Omron CX-Programmer project OmronTeachingExample (CX-Programmer 9.73)

# PLC ExamplePLC: CP1H XA

## Program Main (cyclic task 0)

### Section Section1

### Section Analog_Validity

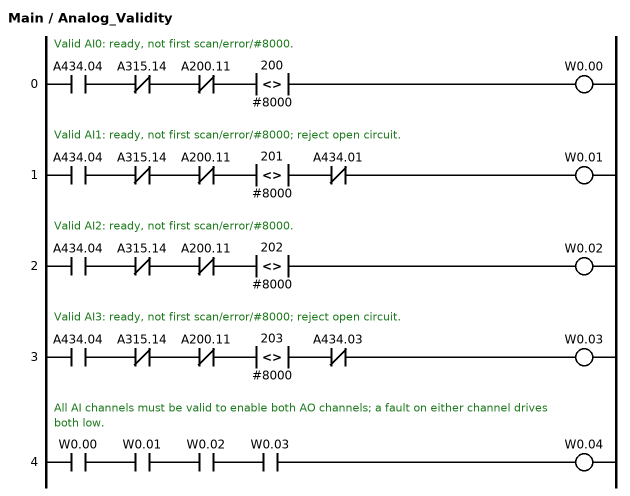
; rung 0: Valid AI0: ready, not first scan/error/#8000.
LD A434.04
ANDNOT A315.14
ANDNOT A200.11
AND<>(305) 200 #8000
OUT W0.00
; rung 1: Valid AI1: ready, not first scan/error/#8000; reject open circuit.
LD A434.04
ANDNOT A315.14
ANDNOT A200.11
AND<>(305) 201 #8000
ANDNOT A434.01
OUT W0.01
; rung 2: Valid AI2: ready, not first scan/error/#8000.
LD A434.04
ANDNOT A315.14
ANDNOT A200.11
AND<>(305) 202 #8000
OUT W0.02
; rung 3: Valid AI3: ready, not first scan/error/#8000; reject open circuit.
LD A434.04
ANDNOT A315.14
ANDNOT A200.11
AND<>(305) 203 #8000
ANDNOT A434.03
OUT W0.03
; rung 4: All AI channels must be valid to enable both AO channels; a fault on either channel drives both low.
LD W0.00
AND W0.01
AND W0.02
AND W0.03
OUT W0.04

### Section HMI_Input_Publication

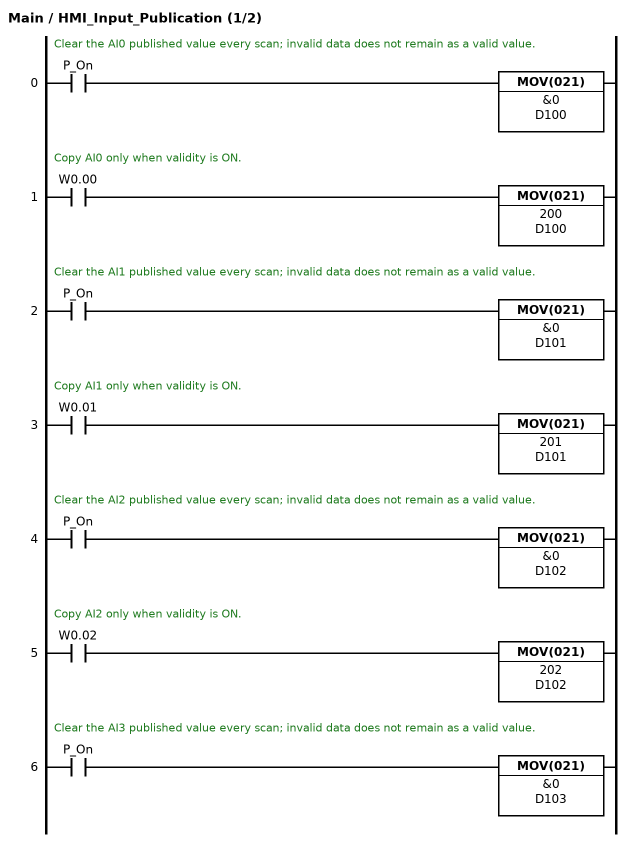
; rung 0: Clear the AI0 published value every scan; invalid data does not remain as a valid value.
LD P_On
MOV(021) &0 D100
; rung 1: Copy AI0 only when validity is ON.
LD W0.00
MOV(021) 200 D100
; rung 2: Clear the AI1 published value every scan; invalid data does not remain as a valid value.
LD P_On
MOV(021) &0 D101
; rung 3: Copy AI1 only when validity is ON.
LD W0.01
MOV(021) 201 D101
; rung 4: Clear the AI2 published value every scan; invalid data does not remain as a valid value.
LD P_On
MOV(021) &0 D102
; rung 5: Copy AI2 only when validity is ON.
LD W0.02
MOV(021) 202 D102
; rung 6: Clear the AI3 published value every scan; invalid data does not remain as a valid value.
LD P_On
MOV(021) &0 D103

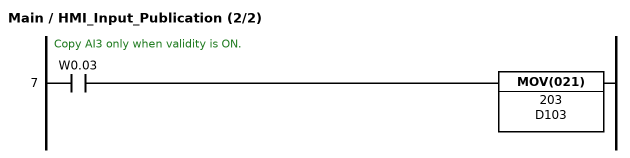
; rung 7: Copy AI3 only when validity is ON.
LD W0.03
MOV(021) 203 D103

### Section AO_Command_Arbitration

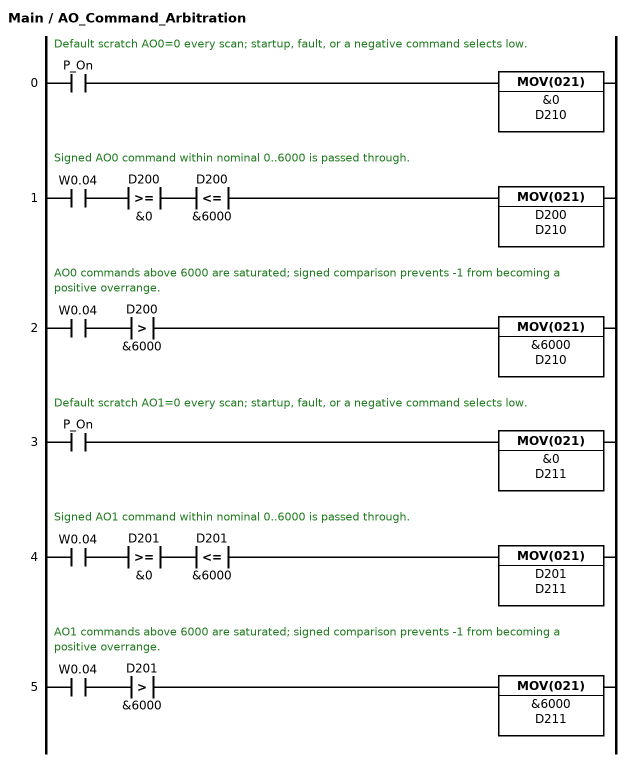
; rung 0: Default scratch AO0=0 every scan; startup, fault, or a negative command selects low.
LD P_On
MOV(021) &0 D210
; rung 1: Signed AO0 command within nominal 0..6000 is passed through.
LD W0.04
AND>=S(327) D200 &0
AND<=S(317) D200 &6000
MOV(021) D200 D210
; rung 2: AO0 commands above 6000 are saturated; signed comparison prevents -1 from becoming a positive overrange.
LD W0.04
AND>S(322) D200 &6000
MOV(021) &6000 D210
; rung 3: Default scratch AO1=0 every scan; startup, fault, or a negative command selects low.
LD P_On
MOV(021) &0 D211
; rung 4: Signed AO1 command within nominal 0..6000 is passed through.
LD W0.04
AND>=S(327) D201 &0
AND<=S(317) D201 &6000
MOV(021) D201 D211
; rung 5: AO1 commands above 6000 are saturated; signed comparison prevents -1 from becoming a positive overrange.
LD W0.04
AND>S(322) D201 &6000
MOV(021) &6000 D211

### Section Final_AO_Writers

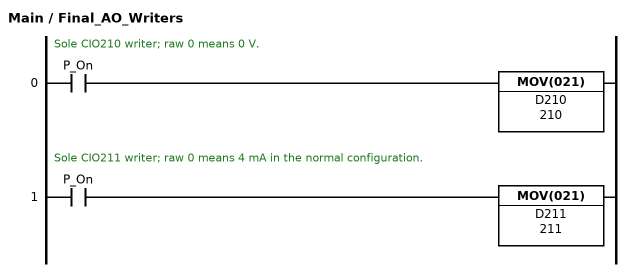
; rung 0: Sole CIO210 writer; raw 0 means 0 V.
LD P_On
MOV(021) D210 210
; rung 1: Sole CIO211 writer; raw 0 means 4 mA in the normal configuration.
LD P_On
MOV(021) D211 211

### Section END
; rung 0
END(001)